FUNCTION F_BuildSelector : STRING
VAR_INPUT
    iValue : UDINT;
END_VAR

F_BuildSelector := CONCAT('00 ', F_UdintToStringPadded(iValue, 2));

END_FUNCTION

(* stored: Version 1.1.0.1
   POU F_BuildSelector: Id {1c9eb3f3-ece6-4d29-baa0-8472cce8052e}, SpecialFunc None *)
